Fanuc KAREL source: ko00054.KL

-- PROVISIONAL review KL for V770-1; original PC SHA256 bc92676fa67a9df99332b3f9adc0c9d2f2775c33cba61ab8961c715bfc03495c
-- Incomplete behavior may be omitted. Consult companion uncertainty JSON. Do not deploy.
PROGRAM KO00054
%NOLOCKGROUP
BEGIN
  -- UNRESOLVED_PC offsets 5-12; opcodes 9D,23
  -- UNRESOLVED_PC offsets 17-69; opcodes 27,27,49,7E,AD,27,49,7E,AD,22,31,7E,4A
  -- UNRESOLVED_PC offsets 74-78; opcodes 7F
END KO00054
